FUNCTION "ROLL_ReadInputs" : Void
{ S7_Optimized_Access := 'TRUE' }
VERSION : 0.1
VAR_TEMP
    b : Int;
    bit : Int;
END_VAR
BEGIN
    // Confirmed four-station profile: absent optional inputs are zero.
    FOR #b := 119 TO 125 DO
        FOR #bit := 0 TO 7 DO "ROLL_IO".Input[#b, #bit] := FALSE; END_FOR;
    END_FOR;
    IF "ROLL_IO".PhysicalIoConfigured AND NOT "ROLL_IO".Simulation THEN
        "ROLL_IO".Input[0, 0] := %I0.0;
        "ROLL_IO".Input[0, 1] := %I0.1;
        "ROLL_IO".Input[0, 2] := %I0.2;
        "ROLL_IO".Input[0, 3] := %I0.3;
        "ROLL_IO".Input[0, 4] := %I0.4;
        "ROLL_IO".Input[0, 5] := %I0.5;
        "ROLL_IO".Input[0, 6] := %I0.6;
        "ROLL_IO".Input[0, 7] := %I0.7;
        "ROLL_IO".Input[1, 0] := %I1.0;
        "ROLL_IO".Input[1, 1] := %I1.1;
        "ROLL_IO".Input[1, 2] := %I1.2;
        "ROLL_IO".Input[1, 3] := %I1.3;
        "ROLL_IO".Input[1, 4] := %I1.4;
        "ROLL_IO".Input[1, 5] := %I1.5;
        "ROLL_IO".Input[1, 6] := %I1.6;
        "ROLL_IO".Input[1, 7] := %I1.7;
        "ROLL_IO".Input[2, 0] := %I2.0;
        "ROLL_IO".Input[2, 1] := %I2.1;
        "ROLL_IO".Input[2, 2] := %I2.2;
        "ROLL_IO".Input[2, 3] := %I2.3;
        "ROLL_IO".Input[2, 4] := %I2.4;
        "ROLL_IO".Input[2, 5] := %I2.5;
        "ROLL_IO".Input[2, 6] := %I2.6;
        "ROLL_IO".Input[2, 7] := %I2.7;
        "ROLL_IO".Input[3, 0] := %I3.0;
        "ROLL_IO".Input[3, 1] := %I3.1;
        "ROLL_IO".Input[3, 2] := %I3.2;
        "ROLL_IO".Input[3, 3] := %I3.3;
        "ROLL_IO".Input[3, 4] := %I3.4;
        "ROLL_IO".Input[3, 5] := %I3.5;
        "ROLL_IO".Input[3, 6] := %I3.6;
        "ROLL_IO".Input[3, 7] := %I3.7;
        "ROLL_IO".Input[4, 0] := %I4.0;
        "ROLL_IO".Input[4, 1] := %I4.1;
        "ROLL_IO".Input[4, 2] := %I4.2;
        "ROLL_IO".Input[4, 3] := %I4.3;
        "ROLL_IO".Input[4, 4] := %I4.4;
        "ROLL_IO".Input[4, 5] := %I4.5;
        "ROLL_IO".Input[4, 6] := %I4.6;
        "ROLL_IO".Input[4, 7] := %I4.7;
        "ROLL_IO".Input[5, 0] := %I5.0;
        "ROLL_IO".Input[5, 1] := %I5.1;
        "ROLL_IO".Input[5, 2] := %I5.2;
        "ROLL_IO".Input[5, 3] := %I5.3;
        "ROLL_IO".Input[5, 4] := %I5.4;
        "ROLL_IO".Input[5, 5] := %I5.5;
        "ROLL_IO".Input[5, 6] := %I5.6;
        "ROLL_IO".Input[5, 7] := %I5.7;
        "ROLL_IO".Input[6, 0] := %I6.0;
        "ROLL_IO".Input[6, 1] := %I6.1;
        "ROLL_IO".Input[6, 2] := %I6.2;
        "ROLL_IO".Input[6, 3] := %I6.3;
        "ROLL_IO".Input[6, 4] := %I6.4;
        "ROLL_IO".Input[6, 5] := %I6.5;
        "ROLL_IO".Input[6, 6] := %I6.6;
        "ROLL_IO".Input[6, 7] := %I6.7;
        "ROLL_IO".Input[7, 0] := %I7.0;
        "ROLL_IO".Input[7, 1] := %I7.1;
        "ROLL_IO".Input[7, 2] := %I7.2;
        "ROLL_IO".Input[7, 3] := %I7.3;
        "ROLL_IO".Input[7, 4] := %I7.4;
        "ROLL_IO".Input[7, 5] := %I7.5;
        "ROLL_IO".Input[7, 6] := %I7.6;
        "ROLL_IO".Input[7, 7] := %I7.7;
        "ROLL_IO".Input[8, 0] := %I8.0;
        "ROLL_IO".Input[8, 1] := %I8.1;
        "ROLL_IO".Input[8, 2] := %I8.2;
        "ROLL_IO".Input[8, 3] := %I8.3;
        "ROLL_IO".Input[8, 4] := %I8.4;
        "ROLL_IO".Input[8, 5] := %I8.5;
        "ROLL_IO".Input[8, 6] := %I8.6;
        "ROLL_IO".Input[8, 7] := %I8.7;
        "ROLL_IO".Input[9, 0] := %I9.0;
        "ROLL_IO".Input[9, 1] := %I9.1;
        "ROLL_IO".Input[9, 2] := %I9.2;
        "ROLL_IO".Input[9, 3] := %I9.3;
        "ROLL_IO".Input[9, 4] := %I9.4;
        "ROLL_IO".Input[9, 5] := %I9.5;
        "ROLL_IO".Input[9, 6] := %I9.6;
        "ROLL_IO".Input[9, 7] := %I9.7;
        "ROLL_IO".Input[10, 0] := %I10.0;
        "ROLL_IO".Input[10, 1] := %I10.1;
        "ROLL_IO".Input[10, 2] := %I10.2;
        "ROLL_IO".Input[10, 3] := %I10.3;
        "ROLL_IO".Input[10, 4] := %I10.4;
        "ROLL_IO".Input[10, 5] := %I10.5;
        "ROLL_IO".Input[10, 6] := %I10.6;
        "ROLL_IO".Input[10, 7] := %I10.7;
        "ROLL_IO".Input[11, 0] := %I11.0;
        "ROLL_IO".Input[11, 1] := %I11.1;
        "ROLL_IO".Input[11, 2] := %I11.2;
        "ROLL_IO".Input[11, 3] := %I11.3;
        "ROLL_IO".Input[11, 4] := %I11.4;
        "ROLL_IO".Input[11, 5] := %I11.5;
        "ROLL_IO".Input[11, 6] := %I11.6;
        "ROLL_IO".Input[11, 7] := %I11.7;
        "ROLL_IO".Input[12, 0] := %I12.0;
        "ROLL_IO".Input[12, 1] := %I12.1;
        "ROLL_IO".Input[12, 2] := %I12.2;
        "ROLL_IO".Input[12, 3] := %I12.3;
        "ROLL_IO".Input[12, 4] := %I12.4;
        "ROLL_IO".Input[12, 5] := %I12.5;
        "ROLL_IO".Input[12, 6] := %I12.6;
        "ROLL_IO".Input[12, 7] := %I12.7;
        "ROLL_IO".Input[13, 0] := %I13.0;
        "ROLL_IO".Input[13, 1] := %I13.1;
        "ROLL_IO".Input[13, 2] := %I13.2;
        "ROLL_IO".Input[13, 3] := %I13.3;
        "ROLL_IO".Input[13, 4] := %I13.4;
        "ROLL_IO".Input[13, 5] := %I13.5;
        "ROLL_IO".Input[13, 6] := %I13.6;
        "ROLL_IO".Input[13, 7] := %I13.7;
        "ROLL_IO".Input[14, 0] := %I14.0;
        "ROLL_IO".Input[14, 1] := %I14.1;
        "ROLL_IO".Input[14, 2] := %I14.2;
        "ROLL_IO".Input[14, 3] := %I14.3;
        "ROLL_IO".Input[14, 4] := %I14.4;
        "ROLL_IO".Input[14, 5] := %I14.5;
        "ROLL_IO".Input[14, 6] := %I14.6;
        "ROLL_IO".Input[14, 7] := %I14.7;
        "ROLL_IO".Input[15, 0] := %I15.0;
        "ROLL_IO".Input[15, 1] := %I15.1;
        "ROLL_IO".Input[15, 2] := %I15.2;
        "ROLL_IO".Input[15, 3] := %I15.3;
        "ROLL_IO".Input[15, 4] := %I15.4;
        "ROLL_IO".Input[15, 5] := %I15.5;
        "ROLL_IO".Input[15, 6] := %I15.6;
        "ROLL_IO".Input[15, 7] := %I15.7;
    END_IF;
END_FUNCTION

FUNCTION "ROLL_WriteOutputs" : Void
{ S7_Optimized_Access := 'TRUE' }
VERSION : 0.1
VAR_TEMP
    enabled : Bool;
END_VAR
BEGIN
    IF "ROLL_IO".PhysicalIoConfigured THEN
        #enabled := "ROLL_IO".PhysicalOutputsEnabled AND NOT "ROLL_IO".Simulation AND NOT "ROLL_IO".ConversionFault;
        %Q16.0 := #enabled AND "ROLL_IO".Output[16, 0];
        %Q16.1 := #enabled AND "ROLL_IO".Output[16, 1];
        %Q16.2 := #enabled AND "ROLL_IO".Output[16, 2];
        %Q16.3 := #enabled AND "ROLL_IO".Output[16, 3];
        %Q16.4 := #enabled AND "ROLL_IO".Output[16, 4];
        %Q16.5 := #enabled AND "ROLL_IO".Output[16, 5];
        %Q16.6 := #enabled AND "ROLL_IO".Output[16, 6];
        %Q16.7 := #enabled AND "ROLL_IO".Output[16, 7];
        %Q17.0 := #enabled AND "ROLL_IO".Output[17, 0];
        %Q17.1 := #enabled AND "ROLL_IO".Output[17, 1];
        %Q17.2 := #enabled AND "ROLL_IO".Output[17, 2];
        %Q17.3 := #enabled AND "ROLL_IO".Output[17, 3];
        %Q17.4 := #enabled AND "ROLL_IO".Output[17, 4];
        %Q17.5 := #enabled AND "ROLL_IO".Output[17, 5];
        %Q17.6 := #enabled AND "ROLL_IO".Output[17, 6];
        %Q17.7 := #enabled AND "ROLL_IO".Output[17, 7];
        %Q18.0 := #enabled AND "ROLL_IO".Output[18, 0];
        %Q18.1 := #enabled AND "ROLL_IO".Output[18, 1];
        %Q18.2 := #enabled AND "ROLL_IO".Output[18, 2];
        %Q18.3 := #enabled AND "ROLL_IO".Output[18, 3];
        %Q18.4 := #enabled AND "ROLL_IO".Output[18, 4];
        %Q18.5 := #enabled AND "ROLL_IO".Output[18, 5];
        %Q18.6 := #enabled AND "ROLL_IO".Output[18, 6];
        %Q18.7 := #enabled AND "ROLL_IO".Output[18, 7];
        %Q19.0 := #enabled AND "ROLL_IO".Output[19, 0];
        %Q19.1 := #enabled AND "ROLL_IO".Output[19, 1];
        %Q19.2 := #enabled AND "ROLL_IO".Output[19, 2];
        %Q19.3 := #enabled AND "ROLL_IO".Output[19, 3];
        %Q19.4 := #enabled AND "ROLL_IO".Output[19, 4];
        %Q19.5 := #enabled AND "ROLL_IO".Output[19, 5];
        %Q19.6 := #enabled AND "ROLL_IO".Output[19, 6];
        %Q19.7 := #enabled AND "ROLL_IO".Output[19, 7];
        %Q20.0 := #enabled AND "ROLL_IO".Output[20, 0];
        %Q20.1 := #enabled AND "ROLL_IO".Output[20, 1];
        %Q20.2 := #enabled AND "ROLL_IO".Output[20, 2];
        %Q20.3 := #enabled AND "ROLL_IO".Output[20, 3];
        %Q20.4 := #enabled AND "ROLL_IO".Output[20, 4];
        %Q20.5 := #enabled AND "ROLL_IO".Output[20, 5];
        %Q20.6 := #enabled AND "ROLL_IO".Output[20, 6];
        %Q20.7 := #enabled AND "ROLL_IO".Output[20, 7];
        %Q21.0 := #enabled AND "ROLL_IO".Output[21, 0];
        %Q21.1 := #enabled AND "ROLL_IO".Output[21, 1];
        %Q21.2 := #enabled AND "ROLL_IO".Output[21, 2];
        %Q21.3 := #enabled AND "ROLL_IO".Output[21, 3];
        %Q21.4 := #enabled AND "ROLL_IO".Output[21, 4];
        %Q21.5 := #enabled AND "ROLL_IO".Output[21, 5];
        %Q21.6 := #enabled AND "ROLL_IO".Output[21, 6];
        %Q21.7 := #enabled AND "ROLL_IO".Output[21, 7];
        %Q22.0 := #enabled AND "ROLL_IO".Output[22, 0];
        %Q22.1 := #enabled AND "ROLL_IO".Output[22, 1];
        %Q22.2 := #enabled AND "ROLL_IO".Output[22, 2];
        %Q22.3 := #enabled AND "ROLL_IO".Output[22, 3];
        %Q22.4 := #enabled AND "ROLL_IO".Output[22, 4];
        %Q22.5 := #enabled AND "ROLL_IO".Output[22, 5];
        %Q22.6 := #enabled AND "ROLL_IO".Output[22, 6];
        %Q22.7 := #enabled AND "ROLL_IO".Output[22, 7];
        %Q23.0 := #enabled AND "ROLL_IO".Output[23, 0];
        %Q23.1 := #enabled AND "ROLL_IO".Output[23, 1];
        %Q23.2 := #enabled AND "ROLL_IO".Output[23, 2];
        %Q23.3 := #enabled AND "ROLL_IO".Output[23, 3];
        %Q23.4 := #enabled AND "ROLL_IO".Output[23, 4];
        %Q23.5 := #enabled AND "ROLL_IO".Output[23, 5];
        %Q23.6 := #enabled AND "ROLL_IO".Output[23, 6];
        %Q23.7 := #enabled AND "ROLL_IO".Output[23, 7];
        %Q24.0 := #enabled AND "ROLL_IO".Output[24, 0];
        %Q24.1 := #enabled AND "ROLL_IO".Output[24, 1];
        %Q24.2 := #enabled AND "ROLL_IO".Output[24, 2];
        %Q24.3 := #enabled AND "ROLL_IO".Output[24, 3];
        %Q24.4 := #enabled AND "ROLL_IO".Output[24, 4];
        %Q24.5 := #enabled AND "ROLL_IO".Output[24, 5];
        %Q24.6 := #enabled AND "ROLL_IO".Output[24, 6];
        %Q24.7 := #enabled AND "ROLL_IO".Output[24, 7];
        %Q25.0 := #enabled AND "ROLL_IO".Output[25, 0];
        %Q25.1 := #enabled AND "ROLL_IO".Output[25, 1];
        %Q25.2 := #enabled AND "ROLL_IO".Output[25, 2];
        %Q25.3 := #enabled AND "ROLL_IO".Output[25, 3];
        %Q25.4 := #enabled AND "ROLL_IO".Output[25, 4];
        %Q25.5 := #enabled AND "ROLL_IO".Output[25, 5];
        %Q25.6 := #enabled AND "ROLL_IO".Output[25, 6];
        %Q25.7 := #enabled AND "ROLL_IO".Output[25, 7];
    END_IF;
END_FUNCTION
